// TIA Portal V20 export
// export: Created 2026-10-19T18:06:42.4107328Z, ExportSetting WithDefaults, DisplayName Totally Integrated Automation Portal, DisplayVersion V20 Update 6, DisplayName TIA Portal Openness, DisplayVersion V20 Update 6, DisplayName TIA Portal Version Control Interface, DisplayVersion V20 Update 6, DisplayName SINAMICS Startdrive Advanced, DisplayVersion V20 SP1, DisplayName SINAMICS Startdrive G130, G150, S120, S150, SINAMICS MV, G220, S200, S210, DisplayVersion V20 SP1, DisplayName SINAMICS Startdrive G110M, G120, G120C, G120D, G120P, G115D, DisplayVersion V20 SP1, DisplayName STEP 7 Professional, DisplayVersion V20 Update 6, DisplayName STEP 7 Safety, DisplayVersion V20 Update 2, DisplayName WinCC Basic/Comfort/Advanced, DisplayVersion V20 Update 6, DisplayName WinCC Unified, DisplayVersion V20 Update 6
DATA_BLOCK "SAI_Cyclic_WeightProc_DB"   // DB29
VERSION : 0.1
// stored: AutoNumber true, DBAccessibleFromOPCUA true, DBAccessibleFromWebserver true, InstanceOfName SAI_Cyclic_WeightProc, InstanceOfType FB
"SAI_Cyclic_WeightProc"
   // VAR_INPUT
   //    WeightCmd { ExternalAccessible := 'False'; ExternalVisible := 'False'; ExternalWritable := 'False'} : Word := 3;
   //    MB_DevStatus : Word;
   // END_VAR
   // VAR_OUTPUT
   //    RealTimeWeight { ExternalVisible := 'False'; ExternalWritable := 'False'} : Real;
   //    StableWeight { ExternalVisible := 'False'; ExternalWritable := 'False'} : Real;
   //    DataOK : Bool;
   //    Motion : Bool;
   //    NetMode : Bool;
   //    Alarm : Bool;
   //    Done { ExternalAccessible := 'False'; ExternalVisible := 'False'; ExternalWritable := 'False'} : Bool;
   //    Error { ExternalAccessible := 'False'; ExternalVisible := 'False'; ExternalWritable := 'False'} : Bool;
   // END_VAR
   // VAR_IN_OUT
   //    TareImmediate { ExternalAccessible := 'False'; ExternalVisible := 'False'; ExternalWritable := 'False'} : Bool;
   //    TareStable { ExternalAccessible := 'False'; ExternalVisible := 'False'; ExternalWritable := 'False'} : Bool;
   //    ZeroImmediate { ExternalAccessible := 'False'; ExternalVisible := 'False'; ExternalWritable := 'False'} : Bool;
   //    ZeroStable { ExternalAccessible := 'False'; ExternalVisible := 'False'; ExternalWritable := 'False'} : Bool;
   //    PreTareValue : Real;
   //    PreTare : Bool;
   //    ClearTare { ExternalAccessible := 'False'; ExternalVisible := 'False'; ExternalWritable := 'False'} : Bool;
   //    MB_Value : Real;
   //    MB_Response : Word;
   //    MB_CmdValue : Real;
   //    MB_Command : Word;
   // END_VAR
   // VAR
   //    WriteTrigger { ExternalAccessible := 'False'; ExternalVisible := 'False'; ExternalWritable := 'False'} : Bool;
   //    RestoreTrigger { ExternalAccessible := 'False'; ExternalVisible := 'False'; ExternalWritable := 'False'} : Bool;
   //    Cmd { ExternalAccessible := 'False'; ExternalVisible := 'False'; ExternalWritable := 'False'} : Int;
   //    TareStablePTrigger : Bool;
   //    ZeroStablePTrigger : Bool;
   //    ZeroImmedTrigger : Bool;
   //    TareImmedTrigger : Bool;
   //    ClearTareTrigger : Bool;
   //    PreTareTrigger : Bool;
   // END_VAR
BEGIN
END_DATA_BLOCK
